{attribute 'Tc2GvlVarNames'}
VAR_GLOBAL
	unLOG_INSTANCE_IDX				:UINT;
END_VAR
VAR_GLOBAL CONSTANT
	sLOG_FILE_PATH					:STRING := '\Hard Disk\Riex\Log\';			(* Login file path *)
	sLOG_FILE_SUFFIX					:STRING := 'log';							(* Suffix of loggin file *)
	unNUM_OF_LOG_VAR					:UINT := 4;								(* Number of logging variables *)
	unLOG_MAX_NO						:UINT := 1;
	unLOG_BEFOR_MAX_NO				:UINT := 10;
	unLOG_DURING_MAX_NO				:UINT := 250;
	unLOG_AFTER_MAX_NO				:UINT := 10;
END_VAR

(* stored: Version 1.1.0.1, ProductVersion 3.1.4024.15
   GVL GVL_Logger: Id {be5f59c2-b99c-4f71-a62f-d32808ea0794} *)
